TYPE E_LightAction :
(
    Toggle,
    TurnOn,
    TurnOff
);
END_TYPE

(* stored: Version 1.1.0.1, ProductVersion 3.1.4026.20
   DUT E_LightAction: Id {D1A10002-0A11-4A11-8A11-000000000002} *)
